(* IEC 61131-3 sources: Repository_IEMA_Test/LMC_PacDrive.device.xml.v3^/Plc Logic.plclogic.xml.v3^/Application.application.xml.v3^/TemplateFullProgrammingFramework/Tools, 3 files *)

(* ---- FC_IsDriveVirtual.fn.st ---- *)
FUNCTION FC_IsDriveVirtual : BOOL
VAR_INPUT
	i_ifDrive	: SystemConfigurationItf.IF_Drive;
END_VAR

VAR_OUTPUT
	q_etDiag	: GD.ET_Diag := GD.ET_Diag.Ok;
	q_etDiagExt	: ET_DiagExt := ET_DiagExt.Ok;
	q_sMsg		: STRING[80];
END_VAR

VAR
	xSuccess						: BOOL;
	ifSercosDeviceIdentification	: SystemConfigurationItf.IF_SercosDeviceIdentification;
END_VAR

IF i_ifDrive = 0 THEN
	q_etDiag	:= GD.ET_Diag.InputParameterInvalid;
	q_etDiagExt	:= ET_DiagExt.DriveInvalid;
	q_sMsg		:= 'FC_IsDriveVirtual: i_ifDrive not set';
ELSE
	xSuccess := __QUERYINTERFACE(i_ifDrive, ifSercosDeviceIdentification);
	IF NOT xSuccess OR ifSercosDeviceIdentification = 0 THEN
		q_etDiag	:= GD.ET_Diag.InputParameterInvalid;
		q_etDiagExt	:= ET_DiagExt.DriveInvalid;
		q_sMsg		:= Standard.CONCAT(i_ifDrive.Name, ' - IF_SercosDeviceIdentification not implemented');
	ELSE
		IF ifSercosDeviceIdentification.WorkingState = 0 THEN	// Drive is virtual
			FC_IsDriveVirtual := TRUE;
		ELSE
			FC_IsDriveVirtual := FALSE;
		END_IF
	END_IF
END_IF

(* ---- FC_ObjectTypeIsMotionAxis.fn.st ---- *)
(* Checks whether the given diObjectType is an object representing a Motion Axis (drive beneath SercosIII bus) *)
FUNCTION FC_ObjectTypeIsMotionAxis : BOOL

VAR_INPUT
	i_udiObjectType: UDINT; (* Type (UDINT) of object to be checked to be a motion axis *)
END_VAR

(* Currently, this implemetation is hacky. We compare the ObjectType to a static list of ObjectTypes known as Motion Drives.
   What we acutlly want is to get the IEC object by LogicalAddress and check whether it fits the interface IF_Drive. But sadly,
   such a function doesn't exist yet *)

IF	i_udiObjectType = SystemInterface.LXM62DxS_TYPE.udiType OR
	i_udiObjectType = SystemInterface.ILM62_TYPE.udiType OR
	i_udiObjectType = SystemInterface.LXM52_TYPE.udiType OR
	i_udiObjectType = SystemInterface.SERCDRV_TYPE.udiType OR
	i_udiObjectType = SystemInterface.LXM52Linear_TYPE.udiType OR
	i_udiObjectType = SystemInterface.LXM62DxSLinear_TYPE.udiType
THEN
   FC_ObjectTypeIsMotionAxis := TRUE;
ELSE
   FC_ObjectTypeIsMotionAxis := FALSE;
END_IF

RETURN;

(* ---- FC_SetDeadTimeCompensation.fn.st ---- *)
FUNCTION FC_SetDeadTimeCompensation : BOOL
VAR_INPUT
	i_stSubModuleInterfaceMain		: AXM.ST_Main;
END_VAR
VAR
(* Init related variables *)
	stLogicalAddressMaster			: SystemConfigurationItf.ST_LogicalAddress;
	lrShaftRefDelay					: LREAL;
	lrPositionDelay					: LREAL;
	diResult						: DINT;

END_VAR

IF i_stSubModuleInterfaceMain.i_ifMaster <> 0 AND i_stSubModuleInterfaceMain.i_ifDrive <> 0 THEN
	stLogicalAddressMaster := i_stSubModuleInterfaceMain.i_ifMaster.stLogicalAddress;
	IF (stLogicalAddressMaster.udiType = SYSTEMINTERFACE.P_ENC_TYPE.udiType) OR			(* Physical encoder *)
		(stLogicalAddressMaster.udiType = SYSTEMINTERFACE.INC_IN_TYPE.udiType) OR		(* Incremental	encoder *)
		(stLogicalAddressMaster.udiType = SYSTEMINTERFACE.V_ENC_TYPE.udiType) THEN		(* Virtual master encoder *)

		stLogicalAddressMaster := i_stSubModuleInterfaceMain.i_ifDrive.stLogicalAddress;
		stLogicalAddressMaster.udiParameterId := 16#00A2;
		diResult := SYSTEMINTERFACE.FC_GetParameter(i_stLogAdr	:= stLogicalAddressMaster,
													i_dwBuffer	:= ADR(lrShaftRefDelay),
													i_diSize	:= SIZEOF(lrShaftRefDelay));
		IF diResult = 0 THEN
			i_stSubModuleInterfaceMain.iq_lencEncoder.Delay := -lrShaftRefDelay;
		END_IF
	ELSIF (stLogicalAddressMaster.udiType = SYSTEMINTERFACE.INC_IN3_TYPE.udiType) THEN  (* IncIn via TM5 TM5SE1IC20005 *)
		stLogicalAddressMaster := i_stSubModuleInterfaceMain.i_ifDrive.stLogicalAddress;
		stLogicalAddressMaster.udiParameterId := 16#00A2;
		diResult := SYSTEMINTERFACE.FC_GetParameter(i_stLogAdr	:= stLogicalAddressMaster,
													i_dwBuffer	:= ADR(lrShaftRefDelay),
													i_diSize	:= SIZEOF(lrShaftRefDelay));
		IF diResult = 0 THEN
			i_stSubModuleInterfaceMain.iq_lencEncoder.Delay := -lrShaftRefDelay;
			stLogicalAddressMaster := i_stSubModuleInterfaceMain.i_ifMaster.stLogicalAddress;
			stLogicalAddressMaster.udiParameterId := 16#008E; 					(* Parameter PositionDelay of TM5SE1IC20005 *)
			diResult := SYSTEMINTERFACE.FC_GetParameter(i_stLogAdr	:= stLogicalAddressMaster,
														i_dwBuffer	:= ADR(lrPositionDelay),
														i_diSize	:= SIZEOF(lrPositionDelay));
			IF diResult = 0 THEN
				i_stSubModuleInterfaceMain.iq_lencEncoder.Delay := -(lrShaftRefDelay + (-lrPositionDelay)) ;
			END_IF
		END_IF
	END_IF
END_IF

IF diResult = 0 THEN
	FC_SetDeadTimeCompensation := TRUE;
END_IF
